Fanuc KAREL source: KB00058.KL

PROGRAM KB00058
%NOLOCKGROUP
VAR
  P1: INTEGER
  P2: STRING[80]
  P3: STRING[80]
  P4: INTEGER
BEGIN
  P1 = 1
  P2 = 'A'
  P3 = 'A'
  P4 = 1
  DAQ_WRITE(P1, P2, P3, P4)
END KB00058
